(* IEC 61131-3 sources: Test-Git_ESME26/TestProgettoESME_26.fbsproj/TemplateFullProgrammingFramework_Migration.device.xml.v3^/Plc Logic.plclogic.xml.v3^/Application.application.xml.v3^/TemplateFullProgrammingFramework/EquipmentModules/SR_AlphaModule.pou.xml.v3^, 7 files *)

(* ---- Init_Master.act.st ---- *)
__METADATA__
{
  "v3Meta": {
    "objectGuid": "5de7a2f5-7513-47c8-ac44-01f3827a8c65",
    "objectTypeGuid": "8ac092e5-3128-4e26-9e7e-11016c6684f2",
    "embeddedObjectTypeGuids": [
      "3b83b776-fb25-43b8-99f2-3c507c9143fc"
    ],
    "properties": {},
    "subObjects": {}
  }
}

(* System generated code, could be modified for your application *)

(* Standard interface *)
astSubModuleInterface[c_udiMaster].i_sModuleName	:= STANDARD.CONCAT(STR1 := iq_stStandardModuleItf.i_sModuleName, STR2 := ': Master');

astSubModuleInterface[c_udiMaster].i_xLogEnable		:= TRUE;
astSubModuleInterface[c_udiMaster].i_wLogDataFilter	:= UDINT_TO_WORD(TPL.ET_LogDataFilter.ModuleDefault);

fbMasterModule.RegisterLoggerPoint(	i_ifParent	:= fbLoggerPoint,
									i_sName		:= 'Master',
									q_etDiag	:= ,
									q_etDiagExt	:= );

(* AxisModule specific interface *)
stMasterInterface.stMain.i_ifMaster		:= i_ifMaster; 		(* Master *)
stMasterInterface.stMain.i_ifDrive		:= DRV_Master.Axis;
stMasterInterface.stMain.iq_lencEncoder	      := LE_Master.Axis;
DRV_Master.Axis.SetAxisTypeModulo(i_lrPeriod := 360.0);
DRV_Master.Axis.SetErrorStopRamp(i_lrDeceleration  := 50_000.0,
						  		 i_lrJerk		   := 500_000.0);

xDriveIsVirtual := FC_IsDriveVirtual(	i_ifDrive	:= stMasterInterface.stMain.i_ifDrive,
										q_etDiag	=> etDiag,
										q_etDiagExt	=> etDiagExt,
										q_sMsg		=> sMsgBuffer);

IF etDiag <> GD.ET_Diag.Ok AND NOT xIsDriveVirtualException THEN
	stIsDriveVirtualException.etDiag 	:= etDiag;
	stIsDriveVirtualException.udiDiagExt:= etDiagExt;
	stIsDriveVirtualException.sDiagExt 	:= FC_EtDiagExtToString(i_etDiagExt := etDiagExt);
	stIsDriveVirtualException.sMsg 		:= sMsgBuffer;
	xIsDriveVirtualException 			:= TRUE;
END_IF

fbExceptionHandler.SetException(i_xExceptionActive	:= xIsDriveVirtualException,
								iq_stException		:= stIsDriveVirtualException,
								iq_stExceptionList	:= iq_stExceptionList);

xInitSuccessful := xInitSuccessful AND NOT xIsDriveVirtualException;
etDiag := GD.ET_Diag.Ok;

stMasterInterface.stMain.i_lrMotionActiveVelLimit						:= 15.0;		(* Limit for max. velocity of astAxisModuleInterface to switch output AxisMove in Units/s *)
stMasterInterface.stMain.i_etMotionActiveVelType  						:= AXM_ET_MotionActiveVelType.RefVelocity;

stMasterInterface.stMain.i_timMasterStop								:= T#1S;
stMasterInterface.stMain.i_xHwLimitPos									:= FALSE;
stMasterInterface.stMain.i_xHwLimitNeg									:= FALSE;

stMasterInterface.stMain.stReducedVelocity.i_xEnableReducedVelocity		:= FALSE;
stMasterInterface.stMain.stReducedVelocity.i_xOnlyLimitCheck			:= FALSE;
stMasterInterface.stMain.stReducedVelocity.i_lrMaxReducedVelocity		:= 50.0;

stMasterInterface.stMain.i_xStart										:= FALSE;

(***************************************************************************************************************************************************************************************************)
(*** Homing ***)
	IF xDriveIsVirtual THEN
		stMasterInterface.stHome.i_etMode := PDL_ET_HomeMode.SetPosAxisPosition;			(* Homing Mode  in case of virtual axis *)
	ELSE
		stMasterInterface.stHome.i_etMode := PDL_ET_HomeMode.PosDirectionPosEdgeSensor;						(* Homing Mode in case of real axis *)
	END_IF

	stMasterInterface.stHome.i_xEnableInitAbsReadPos := FALSE;		(* TRUE : Restores the AxisPosition depending on the stHome.etMode
																			  If stHome.i_etMode is equal to PDL_ET_HomeMode.RestorePosFromAxisEncoder or
																			  to PDL_ET_HomeMode.WriteAxisEncoder, the encoder of the axis is read,
																			  or else the position will be restored from the retain area *)

 	stMasterInterface.stHome.stSetpos.iq_pstRestorePosRetain := ADR(Grp_stRestorePositionAxis1);

	stMasterInterface.stHome.i_xResetHomeOk := FALSE;

	(* Possible modes for homing mode Sensor:
		PDL_ET_HomeMode.PosDirectionPosEdgeSensor
		PDL_ET_HomeMode.NegDirectionPosEdgeSensor
		PDL_ET_HomeMode.NegDirectionNegEdgeSensor
		PDL_ET_HomeMode.PosDirectionNegEdgeSensor
	*)
	stMasterInterface.stHome.stSensor.i_lrHomePosition			:= 0.0;			(* Position at the end of homing in units *)
	stMasterInterface.stHome.stSensor.i_lrVel					:= 10.0;		(* Homing ceiling velocity in units/s *)
	stMasterInterface.stHome.stSensor.i_lrAcc					:= 1000.0;		(* Homing acceleration in units/s^2 *)
	stMasterInterface.stHome.stSensor.i_lrDec					:= 1000.0;		(* Homing deceleration in units/s^2 *)
	stMasterInterface.stHome.stSensor.i_lrJerk					:= 10000.0;		(* Homing jerk in units/s^3 *)
	stMasterInterface.stHome.stSensor.i_lrOffset				:= 0.0;			(* Offset from home signal in units *)
	stMasterInterface.stHome.stSensor.i_lrMaxTravel				:= 720.0;		(* Max. travel for referencing by normal input *)
	stMasterInterface.stHome.stSensor.i_xRotativeSystem			:= FALSE;		(* Rotative system true or false for referencing by normal input *)
	stMasterInterface.stHome.stSensor.i_xSensor					:= FALSE;		(* Input for home signal. Can be a signal from a controller input. Has to be written cyclic. *)

	(* Possible Modes for homing mode LimitSwitch:
		PDL_ET_HomeMode.PosDirectionPosEdgeHWLimitPos		normally open contact / Closing contact
		PDL_ET_HomeMode.NegDirectionPosEdgeHWLimitNeg		normally open contact / Closing contact
		PDL_ET_HomeMode.NegDirectionNegEdgeHWLimitNeg		normally closed contact / Opening contact
		PDL_ET_HomeMode.PosDirectionNegEdgeHWLimitPos		normally closed contact / Opening contact
	*)
	stMasterInterface.stHome.stLimitSwitch.i_lrHomePosition		:= 0.0;			(* Position at the end of homing in units *)
	stMasterInterface.stHome.stLimitSwitch.i_lrVel				:= 10.0;		(* Homing ceiling velocity in units/s *)
	stMasterInterface.stHome.stLimitSwitch.i_lrLowVel			:= 5.0;			(* Homing low ceiling velocity in units/s *)
	stMasterInterface.stHome.stLimitSwitch.i_lrAcc				:= 1000.0;		(* Homing acceleration in units/s^2 *)
	stMasterInterface.stHome.stLimitSwitch.i_lrDec				:= 1000.0;		(* Homing deceleration in units/s^2 *)
	stMasterInterface.stHome.stLimitSwitch.i_lrJerk				:= 10000.0;		(* Homing jerk in units/s^3 *)
	stMasterInterface.stHome.stLimitSwitch.i_lrOffset			:= 0.0;			(* Offset from home signal in units *)
	stMasterInterface.stHome.stLimitSwitch.i_lrMaxTravel		:= 9999.0;		(* Max. travel for referencing normal input as a hardware limit *)

	(* Possible modes for homing mode MoveOnPos:
		PDL_ET_HomeMode.MoveOnPosAbs
	*)
	stMasterInterface.stHome.stMoveOnPos.i_lrTarget				:= 0.0;			(* Position at the end of homing in units *)
	stMasterInterface.stHome.stMoveOnPos.i_lrVel				:= 10.0;		(* Homing ceiling velocity in units/s *)
	stMasterInterface.stHome.stMoveOnPos.i_lrAcc				:= 1000.0;		(* Homing acceleration in units/s^2 *)
	stMasterInterface.stHome.stMoveOnPos.i_lrDec				:= 1000.0;		(* Homing deceleration in units/s^2 *)
	stMasterInterface.stHome.stMoveOnPos.i_lrJerk				:= 10000.0;		(* Homing jerk in units/s^3 *)
	stMasterInterface.stHome.stMoveOnPos.i_lrPeriod				:= 0.0;			(* Period of the axis *)
	stMasterInterface.stHome.stMoveOnPos.i_xRotativeSystem		:= FALSE;		(* Rotative system true or false *)

	(* Possible modes for homing mode SetPos:
		PDL_ET_HomeMode.SetPosAxisPosition
		PDL_ET_HomeMode.SetPosLogEncoderPosition
		PDL_ET_HomeMode.SetPosAxisAndLogEncoderPosition
		PDL_ET_HomeMode.RestorePosFromAxisEncoder
		PDL_ET_HomeMode.RestorePosFromRetain
	*)
	stMasterInterface.stHome.stSetpos.i_lrHomePosition			:= 0.0;			(* Position at the end of homing in units *)
	stMasterInterface.stHome.stSetpos.i_lrEncoderPosition		:= 0.0;			(* Encoder position in units after homing *)
	stMasterInterface.stHome.stSetpos.i_lrAbsEncOffset			:= 100.0;		(* Distance to the jump of axis encoder in units  *)
	stMasterInterface.stHome.stSetpos.i_lrRestoreWindow			:= 180;			(* How far can the drive be away from is correct position *)
	stMasterInterface.stHome.stSetpos.i_lrUserPeriod			:= 360;			(* Period of the axis *)
	stMasterInterface.stHome.stSetPos.i_xKeepPowerDisabled 		:= FALSE;		(* Keep Power disabled during SetPosHoming true or false*)

	(* Possible modes for homing mode Torque:
		PDL_ET_HomeMode.PosDirectionMaxTorque
		PDL_ET_HomeMode.NegDirectionMaxTorque
	*)
	stMasterInterface.stHome.stTorque.i_lrHomePosition			:= 0.0;			(* Position at the end of homing in units *)
	stMasterInterface.stHome.stTorque.i_lrVel					:= 10.0;		(* Homing ceiling velocity in units/s *)
	stMasterInterface.stHome.stTorque.i_lrAcc					:= 1000.0;		(* Homing acceleration in units/s^2 *)
	stMasterInterface.stHome.stTorque.i_lrDec					:= 1000.0;		(* Homing deceleration in units/s^2 *)
	stMasterInterface.stHome.stTorque.i_lrJerk					:= 10000.0;		(* Homing jerk in units/s^3 *)
	stMasterInterface.stHome.stTorque.i_lrOffset				:= 0.0;			(* Offset from home signal in units *)
	stMasterInterface.stHome.stTorque.i_lrMaxTravel				:= 9999.0;		(* Max. travel for referencing by torque *)
	stMasterInterface.stHome.stTorque.i_lrMaxTorque				:= 0.0;			(* Torque for stop in Nm / referencing by torque *)
	stMasterInterface.stHome.stTorque.i_diTorqueTime			:= 5;			(* Time in msec to hold torque *)

	(* Possible modes for homing mode TouchProbe:
		PDL_ET_HomeMode.PosDirectionPosEdgeTp
		PDL_ET_HomeMode.NegDirectionPosEdgeTp
		PDL_ET_HomeMode.NegDirectionNegEdgeTp
		PDL_ET_HomeMode.PosDirectionNegEdgeTp
	*)
	stMasterInterface.stHome.stTouchProbe.i_lrHomePosition		:= 0.0;			(* Position at the end of homing in units *)
	stMasterInterface.stHome.stTouchProbe.i_lrVel				:= 100.0;		(* Homing ceiling velocity in units/s *)
	stMasterInterface.stHome.stTouchProbe.i_lrAcc				:= 1000.0;		(* Homing acceleration in units/s^2 *)
	stMasterInterface.stHome.stTouchProbe.i_lrDec				:= 1000.0;		(* Homing deceleration in units/s^2 *)
	stMasterInterface.stHome.stTouchProbe.i_lrJerk				:= 10000.0;		(* Homing jerk in units/s^3 *)
	stMasterInterface.stHome.stTouchProbe.i_lrOffset			:= 30.0;		(* Offset from home signal in units *)
	stMasterInterface.stHome.stTouchProbe.i_lrMaxTravel			:= 720.0;		(* Max. travel for referencing by TP *)
	stMasterInterface.stHome.stTouchProbe.i_xRotativeSystem		:= TRUE;		(* Rotative system true or false for referencing by TP *)
 	stMasterInterface.stHome.stTouchProbe.i_ifTouchProbe		:= 0;		(* Input for TP *)

	(* Possible modes for homing mode WritePos:
		PDL_ET_HomeMode.WriteAxisEncoder
	*)
	stMasterInterface.stHome.stWritePos.i_lrHomePosition		:= 0.0;			(* Position at the end of homing in units *)
	stMasterInterface.stHome.stWritePos.i_lrUserPeriod			:= 0.0;			(* Calculates Drive.Position into period ( units ) *)
	stMasterInterface.stHome.stWritePos.i_lrAbsEncOffset		:= 100.0;		(* Distance to the jump of axis encoder in units *)
(***************************************************************************************************************************************************************************************************)
(*** Manual ***)
	stMasterInterface.stManual.i_lrVel								:= 50.0;			(* Velocity in units/s *)
	stMasterInterface.stManual.i_lrAcc								:= 100.0;			(* Acceleration in units/s^2 *)
	stMasterInterface.stManual.i_lrDec								:= 100.0;			(* Deceleration in units/s^2 *)
	stMasterInterface.stManual.i_lrJerk								:= 1000.0;			(* Jerk in units/s^3 *)
	stMasterInterface.stManual.i_lrMaxDistance						:= 120.0;			(* Max pathlengths for one step in units *)
	stMasterInterface.stManual.i_xEndless							:= FALSE;			(* TRUE: jogging endless; Position between the periode; FALSE: jogging in steps. Position can be out of periode *)
	stMasterInterface.stManual.i_lrPeriod							:= 360.0;			(* Period of the axis *)

(***************************************************************************************************************************************************************************************************)
(*** Endless ***)
	stMasterInterface.stEndless.i_lrPeriod 				:= 360.0;		(* Period one cycle in units *)
	stMasterInterface.stEndless.i_lrJerk 				:= 108000.0;	(* Jerk in units/s^3 *)
	stMasterInterface.stEndless.i_lrStopPosition 		:= 120.0;		(* Stop position in units *)
	stMasterInterface.stEndless.i_lrAcc  				:= 10800.0;		(* Acceleration in Units/s^2 *)
	stMasterInterface.stEndless.i_lrDec  				:= 10800.0;		(* Deceleration in Units/s^2 *)
	stMasterInterface.stEndless.i_lrVel 				:= 180.0;   	(* Velocity in Units/s *)

(***************************************************************************************************************************************************************************************************)
(*** Pos ***)
	stMasterInterface.stPos.i_etPosMode					:= PDL_ET_PosMode.Relative;		(* SYSTEMINTERFACE.ET_PosMode.Endless, SYSTEMINTERFACE.ET_PosMode.Relative, SYSTEMINTERFACE.ET_PosMode.Absolute *)
	stMasterInterface.stPos.i_lrTarget 					:= 1440.0;		(* Target position or distance in Units *)
	stMasterInterface.stPos.i_lrAcc 					:= 10800.0;		(* Acceleration in Units/s^2 *)
	stMasterInterface.stPos.i_lrDec 					:= 10800.0;		(* Deceleration in Units/s^2 *)
	stMasterInterface.stPos.i_lrJerk 					:= 108000.0;	(* Jerk in units/s^3 *)
	stMasterInterface.stPos.i_lrVel 					:= 540.0;		(* Ceiling velocity in Units/s *)

// stMasterInterface.stPos.i_xStop								:= FALSE;
(* End of system generated code, could be modified for your application *)

(* ---- Init_Reactions.act.st ---- *)
__METADATA__
{
  "v3Meta": {
    "objectGuid": "b8c61856-85d5-4516-9382-6d221f6f28d2",
    "objectTypeGuid": "8ac092e5-3128-4e26-9e7e-11016c6684f2",
    "embeddedObjectTypeGuids": [
      "3b83b776-fb25-43b8-99f2-3c507c9143fc"
    ],
    "properties": {},
    "subObjects": {}
  }
}

(* System generated code, only to be changed by experienced programmers *)
IF c_udiNumberOfSubModules < 1 THEN
	RETURN;
END_IF

(* Change of default reactions only on demand *)
(* Compare SR MainMachine Action Init_Reactions *)

xInitReactionsException := FALSE;

(*****************************************************************************************************************************************************)
(* Init ReactionTranslationMode *)

TPL.FC_InitReactionTranslationMode(	i_udiNumberOfSubModules			:= c_udiNumberOfSubModules,
									i_petReactionTranslationMode	:= ADR(aetReactionTranslationMode),
									q_etDiag						=> etDiag,
									q_etDiagExt						=> etDiagExtTPL);

IF etDiag <> GD.ET_Diag.Ok AND NOT xInitReactionsException THEN
	xInitReactionsException := TRUE;

	stInitReactionsException.sMsg := SE_CTBX.FC_MultiConcat(i_sString1 := 'InitReactionTranslationMode - ',
														i_sString2 := GD.FC_EtDiagToString(i_etDiag := etDiag),
														i_sString3 := ' - ',
														i_sString4 := TPL.FC_EtDiagExtToString(i_etDiagExt := etDiagExtTPL));
END_IF

(*****************************************************************************************************************************************************)
(* Init ReactionTranslationTable *)

TPL.FC_InitReactionTranslationTable(i_udiNumberOfSubModules			:= c_udiNumberOfSubModules,
									i_pstReactionTranslationTable	:= ADR(aastReactionTranslationTable),
									q_etDiag						=> etDiag,
									q_etDiagExt						=> etDiagExtTPL);

IF etDiag <> GD.ET_Diag.Ok AND NOT xInitReactionsException THEN
	xInitReactionsException := TRUE;

	stInitReactionsException.sMsg := SE_CTBX.FC_MultiConcat(i_sString1 := 'InitReactionTranslationTable - ',
														i_sString2 := GD.FC_EtDiagToString(i_etDiag := etDiag),
														i_sString3 := ' - ',
														i_sString4 := TPL.FC_EtDiagExtToString(i_etDiagExt := etDiagExtTPL));
END_IF

(*****************************************************************************************************************************************************)
(* Init ReactionTranslationJobs *)

TPL.FC_InitReactionTranslationJobs( i_udiNumberOfSubModules			:= c_udiNumberOfSubModules,
									i_pstReactionTranslationJobs	:= ADR(astReactionTranslationJobs),
									q_etDiag						=> etDiag,
									q_etDiagExt						=> etDiagExtTPL);

IF etDiag <> GD.ET_Diag.Ok AND NOT xInitReactionsException THEN
	xInitReactionsException := TRUE;

	stInitReactionsException.sMsg := SE_CTBX.FC_MultiConcat(i_sString1 := 'InitReactionTranslationJobs - ',
														i_sString2 := GD.FC_EtDiagToString(i_etDiag := etDiag),
														i_sString3 := ' - ',
														i_sString4 := TPL.FC_EtDiagExtToString(i_etDiagExt := etDiagExtTPL));
END_IF

(*****************************************************************************************************************************************************)
(* Set exception if any exception occurred *)
fbExceptionHandler.SetException(i_xExceptionActive	:= xInitReactionsException,
								iq_stException		:= stInitReactionsException,
								iq_stExceptionList	:= iq_stExceptionList);

xInitSuccessful := xInitSuccessful AND NOT xInitReactionsException;

etDiag := GD.ET_Diag.Ok;
(* End of system generated code, only to be changed by experienced programmers *)

(* ---- Init_SubModules.act.st ---- *)
__METADATA__
{
  "v3Meta": {
    "objectGuid": "1d297d7a-351d-4413-92a7-7626813427e9",
    "objectTypeGuid": "8ac092e5-3128-4e26-9e7e-11016c6684f2",
    "embeddedObjectTypeGuids": [
      "3b83b776-fb25-43b8-99f2-3c507c9143fc"
    ],
    "properties": {},
    "subObjects": {}
  }
}

(* System generated code, could be modified for your application *)

(* Module Group declaration *)

(* aaudiSubModuleGroups[c_udiAlphaGroup1-TPL.GCL.Gc_udiGroupOffset,TPL.ET_Group.Member1]	:= c_udiMaster; *)	(* The c_diMaster is the first element of the group c_diAlphaGroup1 *)
(* aaudiSubModuleGroups[c_udiAlphaGroup1-TPL.GCL.Gc_udiGroupOffset,TPL.ET_Group.Member2]	:= 0;			*)	(* There is no second element of the group c_diAlphaGroup1 *)

(* aaudiSubModuleGroups[c_udiAlphaGroup2-TPL.GCL.Gc_udiGroupOffset,TPL.ET_Group.Member1]	:= 0;			*)	(* There is no first element of the group c_diAlphaGroup2 *)
(* aaudiSubModuleGroups[c_udiAlphaGroup2-TPL.GCL.Gc_udiGroupOffset,TPL.ET_Group.Member2]	:= 0;			*)	(* There is no second element of the group c_diAlphaGroup2 *)

(* End of system generated code, could be modified for your application *)

(* System generated code, do not change without consulting 'Schneider Electric Automation GmbH' - otherwise you risk instability!!!*)
xInitSubModulesException := FALSE;

(*****************************************************************************************************************************************************)
(* Set IDs of SubModules *)

TPL.FC_SetSubModuleIds(	i_udiMainModuleId			:= iq_stStandardModuleItf.i_udiModuleId,
						i_pstSubModulesItf			:= ADR(astSubModuleInterface),
						i_udiNumberOfSubModules		:= c_udiNumberOfSubModules,
						q_etDiag					=> etDiag,
						q_etDiagExt					=> etDiagExtTPL);

IF etDiag <> GD.ET_Diag.Ok AND NOT xInitSubModulesException THEN
	xInitSubModulesException := TRUE;

	stInitSubModulesException.sMsg := SE_CTBX.FC_MultiConcat(	i_sString1 := 'SetSubModuleIds - ',
															i_sString2 := GD.FC_EtDiagToString(i_etDiag := etDiag),
															i_sString3 := ' - ',
															i_sString4 := TPL.FC_EtDiagExtToString(i_etDiagExt := etDiagExtTPL));
END_IF

(*****************************************************************************************************************************************************)
(* Set exception if any exception occurred *)

fbExceptionHandler.SetException(i_xExceptionActive	:= xInitSubModulesException,
								iq_stException		:= stInitSubModulesException,
								iq_stExceptionList	:= iq_stExceptionList);

xInitSuccessful := xInitSuccessful AND NOT xInitSubModulesException;

etDiag := GD.ET_Diag.Ok;
(* End of system generated code, do not change without consulting 'Schneider Electric Automation GmbH' - otherwise you risk instability!!!*)

(* ---- Output_Active.act.st ---- *)
__METADATA__
{
  "v3Meta": {
    "objectGuid": "2a084c55-f6f9-44d2-9bd5-51403e160ba1",
    "objectTypeGuid": "8ac092e5-3128-4e26-9e7e-11016c6684f2",
    "embeddedObjectTypeGuids": [
      "3b83b776-fb25-43b8-99f2-3c507c9143fc"
    ],
    "properties": {},
    "subObjects": {}
  }
}

(* System generated code, only to be changed by experienced programmers *)
IF iq_stStandardModuleItf.q_udiSubModuleInException <> 0 THEN
	iq_stStandardModuleItf.q_etDiag		:= GD.ET_Diag.Ok;
	iq_stStandardModuleItf.q_udiDiagExt	:= ET_DiagExt.SubModuleInException;
	iq_stStandardModuleItf.q_sDiagExt		:= FC_EtDiagExtToString(i_etDiagExt := ET_DiagExt.SubModuleInException);
	iq_stStandardModuleItf.q_sMsg			:= '';
ELSE
	IF etDiagModuleController = GD.ET_Diag.Ok THEN
		iq_stStandardModuleItf.q_etDiag	:= etDiagModuleController;
		iq_stStandardModuleItf.q_sMsg		:= sMsgModuleController;

		CASE etDiagExtModuleController OF
			TPL.ET_DiagExt.DeactivatingSubModules :
				iq_stStandardModuleItf.q_udiDiagExt	:= ET_DiagExt.DeactivatingSubModules;
				iq_stStandardModuleItf.q_sDiagExt		:= FC_EtDiagExtToString(i_etDiagExt := ET_DiagExt.DeactivatingSubModules);
			TPL.ET_DiagExt.Disabled :
				iq_stStandardModuleItf.q_udiDiagExt	:= ET_DiagExt.Disabled;
				iq_stStandardModuleItf.q_sDiagExt		:= FC_EtDiagExtToString(i_etDiagExt := ET_DiagExt.Disabled);
			TPL.ET_DiagExt.ExecuteStep :
				iq_stStandardModuleItf.q_udiDiagExt	:= ET_DiagExt.ExecuteStep;
				iq_stStandardModuleItf.q_sDiagExt		:= FC_EtDiagExtToString(i_etDiagExt := ET_DiagExt.ExecuteStep);
			TPL.ET_DiagExt.Initializing :
				iq_stStandardModuleItf.q_udiDiagExt	:= ET_DiagExt.Initializing;
				iq_stStandardModuleItf.q_sDiagExt		:= FC_EtDiagExtToString(i_etDiagExt := ET_DiagExt.Initializing);
			TPL.ET_DiagExt.WaitAtNegativeStep :
				iq_stStandardModuleItf.q_udiDiagExt	:= ET_DiagExt.WaitAtNegativeStep;
				iq_stStandardModuleItf.q_sDiagExt		:= FC_EtDiagExtToString(i_etDiagExt := ET_DiagExt.WaitAtNegativeStep);
			TPL.ET_DiagExt.WaitCmdsDone :
				iq_stStandardModuleItf.q_udiDiagExt	:= ET_DiagExt.WaitCmdsDone;
				iq_stStandardModuleItf.q_sDiagExt		:= FC_EtDiagExtToString(i_etDiagExt := ET_DiagExt.WaitCmdsDone);
			TPL.ET_DiagExt.WaitForCmd :
				iq_stStandardModuleItf.q_udiDiagExt	:= ET_DiagExt.WaitForCmd;
				iq_stStandardModuleItf.q_sDiagExt		:= FC_EtDiagExtToString(i_etDiagExt := ET_DiagExt.WaitForCmd);
			ELSE
				iq_stStandardModuleItf.q_etDiag		:= GD. ET_Diag.UnexpectedProgramBehavior;
				iq_stStandardModuleItf.q_udiDiagExt	:= ET_DiagExt.UnknownStateModuleController;
				iq_stStandardModuleItf.q_sDiagExt		:= FC_EtDiagExtToString(i_etDiagExt := ET_DiagExt.UnknownStateModuleController);
		END_CASE
	ELSE
		iq_stStandardModuleItf.q_etDiag		:= GD.ET_Diag.DiagActive;
		iq_stStandardModuleItf.q_udiDiagExt	:= ET_DiagExt.ModuleControllerException;
		iq_stStandardModuleItf.q_sDiagExt		:= FC_EtDiagExtToString(i_etDiagExt := ET_DiagExt.ModuleControllerException);
		iq_stStandardModuleItf.q_sMsg			:= SE_CTBX.FC_MultiConcat(	i_sString1 := GD.FC_EtDiagToString(i_etDiag := etDiagModuleController),
																			i_sString2 := ' - ',
																			i_sString3 := TPL.FC_EtDiagExtToString(i_etDiagExt := etDiagExtModuleController),
																			i_sString4 := '');
	END_IF
END_IF

(* End of system generated code, only to be changed by experienced programmers *)

(* ---- RegisterLoggerPoint.meth.st ---- *)
METHOD RegisterLoggerPoint
VAR_INPUT
	i_ifParent	: APL.IF_LoggerPoint;
	i_sName		: STRING[80];
END_VAR
VAR_OUTPUT
	q_etDiag	: GD.ET_Diag := GD.ET_Diag.Ok;
	q_etDiagExt	: ET_DiagExt := ET_DiagExt.Ok;
END_VAR

fbLoggerPoint.RegisterLoggerPoint(	i_ifParent	:= i_ifParent,
									i_sName		:= i_sName,
									i_sType		:= 'Node Module',
									i_sSource	:= 'Program',
									q_etDiag	=> ,
									q_etDiagExt	=> );

(* ---- Start_Action.act.st ---- *)
__METADATA__
{
  "v3Meta": {
    "objectGuid": "4cbd4b3c-7bad-4b2b-8753-f3e45c041021",
    "objectTypeGuid": "8ac092e5-3128-4e26-9e7e-11016c6684f2",
    "embeddedObjectTypeGuids": [
      "3b83b776-fb25-43b8-99f2-3c507c9143fc"
    ],
    "properties": {},
    "subObjects": {}
  }
}

(* This step is active until the machine is being enabled *)

(* System generated code, do not change without consulting 'Schneider Electric Automation GmbH' - otherwise you risk instability!!! *)
iq_stStandardModuleItf.q_xActive			:= FALSE;
iq_stStandardModuleItf.q_xReady				:= FALSE;

iq_stStandardModuleItf.q_etDiag				:= GD.ET_Diag.Ok;
iq_stStandardModuleItf.q_udiDiagExt			:= ET_DiagExt.Disabled;
iq_stStandardModuleItf.q_sDiagExt			:= FC_EtDiagExtToString(i_etDiagExt := iq_stStandardModuleItf.q_udiDiagExt);
iq_stStandardModuleItf.q_sMsg				:= '';

iq_stStandardModuleItf.q_dwModuleType		:= TPL.ET_ModuleType.NodeModule;
iq_stStandardModuleItf.q_sModuleTypeName	:= 'NodeModule';
iq_stStandardModuleItf.q_udiModuleVersion	:= 1;
(* End of system generated code, do not change without consulting 'Schneider Electric Automation GmbH' - otherwise you risk instability!!! *)

(* System generated code, to be changed by experienced programmers *)
IF iq_stStandardModuleItf.iq_diCmd <> 0 AND NOT iq_stStandardModuleItf.i_xEnable THEN
	iq_stStandardModuleItf.iq_diCmd := 0;
END_IF
(* End of system generated code, to be changed by experienced programmers *)

(* Application specific code *)
(* ToDo: Add your application specific code here *)
;
(* End of application specific code *)

(* ---- UpdateStructs.act.st ---- *)
__METADATA__
{
  "v3Meta": {
    "objectGuid": "04ac7aa9-2e01-4764-9b60-ec4c0ca11f2c",
    "objectTypeGuid": "8ac092e5-3128-4e26-9e7e-11016c6684f2",
    "embeddedObjectTypeGuids": [
      "3b83b776-fb25-43b8-99f2-3c507c9143fc"
    ],
    "properties": {},
    "subObjects": {}
  }
}

(* System generated code, do not change without consulting 'Schneider Electric Automation GmbH' - otherwise you risk instability!!! *)
fbDetectOnlineChange(	i_xEnable	:= TRUE,
						i_xDetect	:= TRUE,
						q_xActive	=> xDetectOnlineChangeActive,
						q_xReady	=> xDetectOnlineChangeReady,
						q_etDiag	=> etDetectOnlineChangeDiag,
						q_etDiagExt	=> etDetectOnlineChangeDiagExt,
						q_sMsg		=> sDetectOnlineChangeMsg,
						q_xChange	=> );

IF(NOT fbDetectOnlineChange.q_xChange) THEN
	RETURN;
END_IF

iq_stStandardModuleItf.iq_stExt.udiNumberOfSubModules 		:= c_udiNumberOfSubModules;
iq_stStandardModuleItf.iq_stExt.dwSubModulesItf		 		:= ADR(astSubModuleInterface);
iq_stStandardModuleItf.iq_stExt.pdwSubModulesAddItf		 	:= ADR(adwSubModuleAddInterfaces);
iq_stStandardModuleItf.iq_stExt.pstListOfCmdTables			:= ADR(astListOfCmdTables);
iq_stStandardModuleItf.iq_stExt.udiNumberOfCmdTables		:= c_udiNumberOfCmdTables;
(* End of system generated code, do not change without consulting 'Schneider Electric Automation GmbH' - otherwise you risk instability!!! *)

(* System generated code, could be modified for your application *)
xUpdateStructsException := FALSE;

(*****************************************************************************************************************************************************)
(* Update CmdTable - Prepare *)

TPL.FC_UpdateCmdTableListElement(	i_pstListofCmdTables	:= ADR(astListOfCmdTables),
									i_udiNumberOfCmdTables	:= c_udiNumberOfCmdTables,
									i_diCmd					:= ET_Cmd.Prepare,
									i_pstCmdTable			:= ADR(astPrepareTable),
									q_etDiag				=> etDiag,
									q_etDiagExt				=> etDiagExtTPL);

IF etDiag <> GD.ET_Diag.Ok AND NOT xUpdateStructsException THEN
	xUpdateStructsException := TRUE;

	stUpdateStructsException.sMsg := SE_CTBX.FC_MultiConcat(i_sString1 := 'Update CmdTable: Prepare - ',
														i_sString2 := GD.FC_EtDiagToString(i_etDiag := etDiag),
														i_sString3 := ' - ',
														i_sString4 := TPL.FC_EtDiagExtToString(i_etDiagExt := etDiagExtTPL));
END_IF

(*****************************************************************************************************************************************************)
(* Update CmdTable - Auto *)

TPL.FC_UpdateCmdTableListElement(	i_pstListofCmdTables	:= ADR(astListOfCmdTables),
									i_udiNumberOfCmdTables	:= c_udiNumberOfCmdTables,
									i_diCmd					:= ET_Cmd.Auto,
									i_pstCmdTable			:= ADR(astAutoTable),
									q_etDiag				=> etDiag,
									q_etDiagExt				=> etDiagExtTPL);

IF etDiag <> GD.ET_Diag.Ok AND NOT xUpdateStructsException THEN
	xUpdateStructsException := TRUE;

	stUpdateStructsException.sMsg := SE_CTBX.FC_MultiConcat(i_sString1 := 'Update CmdTable: Auto - ',
														i_sString2 := GD.FC_EtDiagToString(i_etDiag := etDiag),
														i_sString3 := ' - ',
														i_sString4 := TPL.FC_EtDiagExtToString(i_etDiagExt := etDiagExtTPL));
END_IF

(*****************************************************************************************************************************************************)
(* Update CmdTable - Manual *)

TPL.FC_UpdateCmdTableListElement(	i_pstListofCMDTables	:= ADR(astListofCMDTables),
									i_udiNumberOfCMDTables	:= c_udiNumberOfCMDTables,
									i_diCMD					:= ET_Cmd.Manual,
									i_pstCMDTable			:= ADR(astManualTable),
									q_etDiag				=> etDiag,
									q_etDiagExt				=> etDiagExtTPL);

IF etDiag <> GD.ET_Diag.Ok AND NOT xUpdateStructsException THEN
	xUpdateStructsException := TRUE;

	stUpdateStructsException.sMsg := SE_CTBX.FC_MultiConcat(i_sString1 := 'Update CmdTable: Manual - ',
														i_sString2 := GD.FC_EtDiagToString(i_etDiag := etDiag),
														i_sString3 := ' - ',
														i_sString4 := TPL.FC_EtDiagExtToString(i_etDiagExt := etDiagExtTPL));
END_IF

(*****************************************************************************************************************************************************)
(* Update CmdTable - Stop *)

TPL.FC_UpdateCmdTableListElement(	i_pstListofCMDTables	:= ADR(astListofCMDTables),
									i_udiNumberOfCMDTables	:= c_udiNumberOfCMDTables,
									i_diCMD					:= ET_Cmd.Stop,
									i_pstCMDTable			:= ADR(astStopTable),
									q_etDiag				=> etDiag,
									q_etDiagExt				=> etDiagExtTPL);

IF etDiag <> GD.ET_Diag.Ok AND NOT xUpdateStructsException THEN
	xUpdateStructsException := TRUE;

	stUpdateStructsException.sMsg := SE_CTBX.FC_MultiConcat(i_sString1 := 'Update CmdTable: Stop - ',
														i_sString2 := GD.FC_EtDiagToString(i_etDiag := etDiag),
														i_sString3 := ' - ',
														i_sString4 := TPL.FC_EtDiagExtToString(i_etDiagExt := etDiagExtTPL));
END_IF

(*****************************************************************************************************************************************************)
(* Update CmdTable - Start *)

TPL.FC_UpdateCmdTableListElement(	i_pstListofCMDTables	:= ADR(astListofCMDTables),
									i_udiNumberOfCmdTables	:= c_udiNumberOfCMDTables,
									i_diCMD					:= ET_Cmd.Start,
									i_pstCMDTable			:= ADR(astStartTable),
									q_etDiag				=> etDiag,
									q_etDiagExt				=> etDiagExtTPL);

IF etDiag <> GD.ET_Diag.Ok AND NOT xUpdateStructsException THEN
	xUpdateStructsException := TRUE;

	stUpdateStructsException.sMsg := SE_CTBX.FC_MultiConcat(i_sString1 := 'Update CmdTable: Start - ',
														i_sString2 := GD.FC_EtDiagToString(i_etDiag := etDiag),
														i_sString3 := ' - ',
														i_sString4 := TPL.FC_EtDiagExtToString(i_etDiagExt := etDiagExtTPL));
END_IF

(*****************************************************************************************************************************************************)
(* Update CmdTable - Abort *)

TPL.FC_UpdateCmdTableListElement(	i_pstListofCMDTables	:= ADR(astListofCMDTables),
									i_udiNumberOfCmdTables	:= c_udiNumberOfCmdTables,
									i_diCMD					:= ET_Cmd.Abort,
									i_pstCMDTable			:= ADR(astAbortTable),
									q_etDiag				=> etDiag,
									q_etDiagExt				=> etDiagExtTPL);

IF etDiag <> GD.ET_Diag.Ok AND NOT xUpdateStructsException THEN
	xUpdateStructsException := TRUE;

	stUpdateStructsException.sMsg := SE_CTBX.FC_MultiConcat(i_sString1 := 'Update CmdTable: Abort - ',
														i_sString2 := GD.FC_EtDiagToString(i_etDiag := etDiag),
														i_sString3 := ' - ',
														i_sString4 := TPL.FC_EtDiagExtToString(i_etDiagExt := etDiagExtTPL));
END_IF

(*****************************************************************************************************************************************************)
(* Update CmdTable - Hold *)

TPL.FC_UpdateCmdTableListElement(	i_pstListofCMDTables	:= ADR(astListofCMDTables),
									i_udiNumberOfCmdTables	:= c_udiNumberOfCmdTables,
									i_diCMD					:= ET_Cmd.Hold,
									i_pstCMDTable			:= ADR(astHoldTable),
									q_etDiag				=> etDiag,
									q_etDiagExt				=> etDiagExtTPL);

IF etDiag <> GD.ET_Diag.Ok AND NOT xUpdateStructsException THEN
	xUpdateStructsException := TRUE;

	stUpdateStructsException.sMsg := SE_CTBX.FC_MultiConcat(i_sString1 := 'Update CmdTable: Hold - ',
														i_sString2 := GD.FC_EtDiagToString(i_etDiag := etDiag),
														i_sString3 := ' - ',
														i_sString4 := TPL.FC_EtDiagExtToString(i_etDiagExt := etDiagExtTPL));
END_IF

(*****************************************************************************************************************************************************)
(* Update CmdTable - BrakeRelease *)

TPL.FC_UpdateCmdTableListElement(	i_pstListofCMDTables	:= ADR(astListofCMDTables),
									i_udiNumberOfCMDTables	:= c_udiNumberOfCMDTables,
									i_diCMD					:= ET_Cmd.BrakeRelease,
									i_pstCMDTable			:= ADR(astBrakeReleaseTable),
									q_etDiag				=> etDiag,
									q_etDiagExt				=> etDiagExtTPL);

IF etDiag <> GD.ET_Diag.Ok AND NOT xUpdateStructsException THEN
	xUpdateStructsException := TRUE;

	stUpdateStructsException.sMsg := SE_CTBX.FC_MultiConcat(i_sString1 := 'Update CmdTable: BrakeRelease - ',
														i_sString2 := GD.FC_EtDiagToString(i_etDiag := etDiag),
														i_sString3 := ' - ',
														i_sString4 := TPL.FC_EtDiagExtToString(i_etDiagExt := etDiagExtTPL));
END_IF

(*****************************************************************************************************************************************************)
(* Update AddInterface - Master *)

AXM_FC_UpdateAddInterfaceStruct(	i_pdwSubModuleAddInterfaces	:= ADR(adwSubModuleAddInterfaces),
									i_udiSubModuleConstant		:= c_udiMaster,
									iq_stAxisModuleItf			:= stMasterInterface,
									q_etDiag					=> etDiag,
									q_etDiagExt					=> etDiagExtAXM);

IF etDiag <> GD.ET_Diag.Ok AND NOT xUpdateStructsException THEN
	xUpdateStructsException := TRUE;

	stUpdateStructsException.sMsg := SE_CTBX.FC_MultiConcat(i_sString1 := 'Update AddInterface: Master - ',
														i_sString2 := GD.FC_EtDiagToString(i_etDiag := etDiag),
														i_sString3 := ' - ',
														i_sString4 := AXM_FC_EtDiagExtToString(i_etDiagExt := etDiagExtAXM));
END_IF

(*****************************************************************************************************************************************************)
(* Update ILS Data *)

// stMasterInterface.stEndless.pstIlsData	:= ADR(G_stIlsData);
// stMasterInterface.stMultiCam.pstIlsData	:= ADR(G_stIlsData);

(*****************************************************************************************************************************************************)
(* Set exception if any exception occurred *)

fbExceptionHandler.SetException(i_xExceptionActive	:= xUpdateStructsException,
								iq_stException		:= stUpdateStructsException,
								iq_stExceptionList	:= iq_stExceptionList);

xInitSuccessful := xInitSuccessful AND NOT xUpdateStructsException;

etDiag := GD.ET_Diag.Ok;
(* End of system generated code, could be modified for your application *)
